(* IEC 61131-3 sources: codesys-to-s7/tests/corpus/C2S7-ADDR-MAP/pos, 1 file *)

(* ---- input.st ---- *)
VAR_GLOBAL
    xIn AT %IX0.3 : BOOL;
    iRaw AT %IW5 : INT;
END_VAR
